(* PLC project , CODESYS CODESYS V3.5 SP16 Patch 4 *)
(* stored: creationDateTime 2021-05-05T17:31:41.2561045, modificationDateTime 2021-05-05T17:31:08.0878849 *)

FUNCTION_BLOCK trip_logic
  VAR_INPUT
    PV_OUT : INT;
    TSP : INT;
    TRIP_LOGIC : BOOL;
    K_DELAY : TIME;
  END_VAR
  VAR_OUTPUT
    TRIP_LOGIC_out : BOOL;
    TON1_ET : TIME;
  END_VAR
  VAR
    TON_0 : TON;
  END_VAR

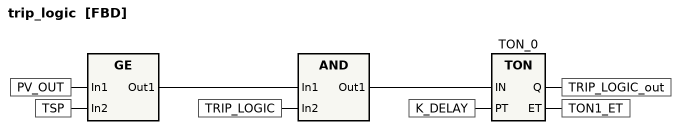
(* FBD diagram, written out as Structured Text *)
TON_0(IN := PV_OUT >= TSP AND TRIP_LOGIC, PT := K_DELAY, ET => TON1_ET);
TRIP_LOGIC_out := TON_0.Q;
END_FUNCTION_BLOCK
